(* IEC 61131-3 sources: nautilus/cmd/naut/testdata/snmp, 1 file *)

(* ---- hw_types.st ---- *)
(*
  Generated by `naut snmp import`: the IT-hardware UDT set from
  docs/design/it-drivers.md §2. Do not edit — every importer (snmp, redfish,
  prometheus) writes this same file, so re-running any of them restores it.
  Member order is the wire order the drivers deliver; the compiled TYPE
  must match it slot for slot, which is why it is generated and not typed.
*)

TYPE
  CPU : STRUCT
    Model : STRING;
    Cores : DINT;
    Health : DINT;
    Fault : BOOL;
    TempC : REAL;
    Pct : REAL;
  END_STRUCT;
  CephCluster : STRUCT
    Online : BOOL;
    HealthStatus : DINT;
    HealthOK : BOOL;
    Fault : BOOL;
    Warning : BOOL;
    OsdTotal : DINT;
    OsdUp : DINT;
    OsdIn : DINT;
    MonQuorum : DINT;
    MgrActive : BOOL;
    PgDegraded : DINT;
    ObjectsDegraded : DINT;
    UsedPct : REAL;
  END_STRUCT;
  CnpgCluster : STRUCT
    Online : BOOL;
    Instances : DINT;
    Primaries : DINT;
    Primary : STRING;
    StreamingReplicas : DINT;
    LagS : REAL;
    BackupAgeS : REAL;
    Fault : BOOL;
  END_STRUCT;
  DIMM : STRUCT
    Locator : STRING;
    CapacityGB : REAL;
    Manufacturer : STRING;
    PartNumber : STRING;
    Health : DINT;
    Fault : BOOL;
    TempC : REAL;
  END_STRUCT;
  Drive : STRUCT
    Bay : DINT;
    Name : STRING;
    Model : STRING;
    Serial : STRING;
    CapacityGB : REAL;
    Protocol : STRING;
    MediaType : STRING;
    Health : DINT;
    Fault : BOOL;
    PredictedFailure : BOOL;
    TempC : REAL;
    Present : BOOL;
  END_STRUCT;
  ErpsRing : STRUCT
    Online : BOOL;
    Idle : BOOL;
    SignalFail : BOOL;
    RplBlocked : BOOL;
    PortsForwarding : DINT;
    Members : DINT;
    FactsAgeS : REAL;
    Stale : BOOL;
    Fault : BOOL;
  END_STRUCT;
  Fan : STRUCT
    Name : STRING;
    Present : BOOL;
    RPM : REAL;
    Pct : REAL;
    Fault : BOOL;
  END_STRUCT;
  IncusCluster : STRUCT
    Online : BOOL;
    MembersTotal : DINT;
    MembersOnline : DINT;
    HealingThreshold : DINT;
    InstancesRunning : DINT;
    Fault : BOOL;
  END_STRUCT;
  KubeCluster : STRUCT
    Online : BOOL;
    NodesTotal : DINT;
    NodesReady : DINT;
    Fault : BOOL;
  END_STRUCT;
  NetPort : STRUCT
    Name : STRING;
    LinkUp : BOOL;
    SpeedGbps : REAL;
    MAC : STRING;
  END_STRUCT;
  PCIeDevice : STRUCT
    Slot : DINT;
    Name : STRING;
    Model : STRING;
    Manufacturer : STRING;
    Firmware : STRING;
    Health : DINT;
    Fault : BOOL;
    Ports : DINT;
    TempC : REAL;
  END_STRUCT;
  PDU : STRUCT
    Online : BOOL;
    Name : STRING;
    Model : STRING;
    Serial : STRING;
    Amps : REAL;
    Watts : REAL;
    Overload : BOOL;
    OutletCount : DINT;
  END_STRUCT;
  PDUOutlet : STRUCT
    Index : DINT;
    Name : STRING;
    On : BOOL;
    Amps : REAL;
    Watts : REAL;
  END_STRUCT;
  PSU : STRUCT
    Name : STRING;
    Present : BOOL;
    Fault : BOOL;
    InputOk : BOOL;
    InputV : REAL;
    OutputW : REAL;
    CapacityW : REAL;
  END_STRUCT;
  Probe : STRUCT
    Online : BOOL;
    Kind : STRING;
    Target : STRING;
    Up : BOOL;
    DurationS : REAL;
    HttpStatus : DINT;
    Expected : STRING;
    Fault : BOOL;
  END_STRUCT;
  PromAlerts : STRUCT
    Firing : DINT;
    Critical : DINT;
    Warning : DINT;
    AnyCritical : BOOL;
    AnyWarning : BOOL;
    Worst : STRING;
  END_STRUCT;
  Server : STRUCT
    Online : BOOL;
    PowerOn : BOOL;
    Health : DINT;
    Fault : BOOL;
    Warning : BOOL;
    Model : STRING;
    Serial : STRING;
    UptimeS : DINT;
    CpuPct : REAL;
    MemPct : REAL;
    Load1 : REAL;
    RootDiskPct : REAL;
    InletTempC : REAL;
    MaxTempC : REAL;
    PowerW : REAL;
    FanCount : DINT;
    PsuCount : DINT;
    TempCount : DINT;
  END_STRUCT;
  Switch : STRUCT
    Online : BOOL;
    Name : STRING;
    Model : STRING;
    Serial : STRING;
    UptimeS : DINT;
    CpuPct : REAL;
    MemPct : REAL;
    TempC : REAL;
    Fault : BOOL;
    PortsTotal : DINT;
    PortsUp : DINT;
  END_STRUCT;
  SwitchPort : STRUCT
    Index : DINT;
    Name : STRING;
    Alias : STRING;
    AdminUp : BOOL;
    OperUp : BOOL;
    Down : BOOL;
    SpeedMbps : REAL;
    InBps : REAL;
    OutBps : REAL;
    InPct : REAL;
    OutPct : REAL;
    InErrors : DINT;
    OutErrors : DINT;
    InDiscards : DINT;
    OutDiscards : DINT;
    ErrorRate : REAL;
    PoeOn : BOOL;
    PoeW : REAL;
    InBroadcastPps : REAL;
    InMulticastPps : REAL;
    Pvid : DINT;
    DiscardRate : REAL;
  END_STRUCT;
  TempSensor : STRUCT
    Name : STRING;
    Value : REAL;
    Fault : BOOL;
    High : BOOL;
    HighHigh : BOOL;
    HighSP : REAL;
    HighHighSP : REAL;
  END_STRUCT;
  UPS : STRUCT
    Online : BOOL;
    Name : STRING;
    Model : STRING;
    Serial : STRING;
    OnBattery : BOOL;
    LowBattery : BOOL;
    BatteryFault : BOOL;
    Fault : BOOL;
    ChargePct : REAL;
    RuntimeMin : REAL;
    LoadPct : REAL;
    InputV : REAL;
    OutputV : REAL;
    BatteryTempC : REAL;
  END_STRUCT;
  VM : STRUCT
    Online : BOOL;
    Present : BOOL;
    Running : BOOL;
    Host : STRING;
    Hosts : DINT;
    Missing : BOOL;
    Conflict : BOOL;
    Expected : STRING;
    Unexpected : BOOL;
    Prefer : STRING;
    Displaced : BOOL;
    OS : STRING;
    CpuPct : REAL;
    MemPct : REAL;
    RootDiskPct : REAL;
    UptimeS : DINT;
    ClockOffsetS : REAL;
    ServicesDown : DINT;
    Fault : BOOL;
  END_STRUCT;
  Vlan : STRUCT
    Id : DINT;
    Name : STRING;
    Ports : STRING;
    Untagged : STRING;
  END_STRUCT;
END_TYPE
